Fanuc KAREL source: kt00959.KL

-- PROVISIONAL review KL for V770-1; original PC SHA256 e95dcc38296ea4a2a5a04b3d77c6f5398ce24e3e879b1d956faf7824ab229719
-- Incomplete behavior may be omitted. Consult companion uncertainty JSON. Do not deploy.
PROGRAM KT00959
%NOLOCKGROUP
VAR
  ENTRY : INTEGER
  PNAME : STRING[80]
  VNAME : STRING[80]
  STATUS : INTEGER
  VALUE : STRING[80]
BEGIN
  -- UNRESOLVED_PC offsets 5-12; opcodes 9C,23
  -- UNRESOLVED_PC offsets 17-25; opcodes 3F,75
  -- UNRESOLVED_PC offsets 30-43; opcodes 3F,75
  -- UNRESOLVED_PC offsets 48-88; opcodes 27,22,22,2A,22,2A,22,2A,22,B0
  -- UNRESOLVED_PC offsets 93-97; opcodes 7F
END KT00959
